{attribute 'qualified_only'}
VAR_GLOBAL
    gAxisConveyor : AXIS_REF;
    gAxisCutter : AXIS_REF;
END_VAR

(* stored: Version 1.1.0.1, ProductVersion 3.1.4024.16
   GVL GVL_Motion: Id {b136a9d1-1841-4446-a6b1-676b2db231e6} *)
